(* IEC 61131-3 sources: llm-plc-st-eval/data/processed_v2/gpt-4o/I3/few_shot, 3 files *)

(* ---- ejec_1.st ---- *)
FUNCTION_BLOCK FB_Alarmas
VAR_INPUT
    alm1 : BOOL; (* Alarma 1 - Prioridad alta *)
    alm2 : BOOL; (* Alarma 2 - Prioridad media *)
    alm3 : BOOL; (* Alarma 3 - Prioridad baja *)
    ack1 : BOOL; (* Reconocimiento de alarma 1 *)
    ack2 : BOOL; (* Reconocimiento de alarma 2 *)
    ack3 : BOOL; (* Reconocimiento de alarma 3 *)
END_VAR
VAR_OUTPUT
    sirena : BOOL; (* Sirena de alarma *)
    codigoAlm : INT; (* Código de la alarma de mayor prioridad *)
END_VAR
VAR
    retAlm1 : BOOL; (* Retención de alarma 1 *)
    retAlm2 : BOOL; (* Retención de alarma 2 *)
    retAlm3 : BOOL; (* Retención de alarma 3 *)
END_VAR

(* Retención de alarmas *)
IF alm1 THEN
    retAlm1 := TRUE;
ELSIF ack1 AND NOT alm1 THEN
    retAlm1 := FALSE;
END_IF;

IF alm2 THEN
    retAlm2 := TRUE;
ELSIF ack2 AND NOT alm2 THEN
    retAlm2 := FALSE;
END_IF;

IF alm3 THEN
    retAlm3 := TRUE;
ELSIF ack3 AND NOT alm3 THEN
    retAlm3 := FALSE;
END_IF;

(* Determinación del código de alarma de mayor prioridad *)
IF retAlm1 THEN
    codigoAlm := 1;
ELSIF retAlm2 THEN
    codigoAlm := 2;
ELSIF retAlm3 THEN
    codigoAlm := 3;
ELSE
    codigoAlm := 0;
END_IF;

(* Activación de la sirena si hay cualquier alarma activa *)
sirena := retAlm1 OR retAlm2 OR retAlm3;

END_FUNCTION_BLOCK

(* ---- ejec_2.st ---- *)
FUNCTION_BLOCK FB_Alarmas
VAR_INPUT
    alm1 : BOOL; (* Alarma 1 - Alta prioridad *)
    alm2 : BOOL; (* Alarma 2 - Media prioridad *)
    alm3 : BOOL; (* Alarma 3 - Baja prioridad *)
    ack1 : BOOL; (* Reconocimiento de alarma 1 *)
    ack2 : BOOL; (* Reconocimiento de alarma 2 *)
    ack3 : BOOL; (* Reconocimiento de alarma 3 *)
END_VAR
VAR_OUTPUT
    sirena : BOOL; (* Sirena de alarma *)
    codigoAlm : INT; (* Código de alarma de mayor prioridad *)
END_VAR
VAR
    retAlm1 : BOOL; (* Retención de alarma 1 *)
    retAlm2 : BOOL; (* Retención de alarma 2 *)
    retAlm3 : BOOL; (* Retención de alarma 3 *)
END_VAR

(* Retención de alarmas *)
IF alm1 THEN
    retAlm1 := TRUE;
ELSIF ack1 AND NOT alm1 THEN
    retAlm1 := FALSE;
END_IF;

IF alm2 THEN
    retAlm2 := TRUE;
ELSIF ack2 AND NOT alm2 THEN
    retAlm2 := FALSE;
END_IF;

IF alm3 THEN
    retAlm3 := TRUE;
ELSIF ack3 AND NOT alm3 THEN
    retAlm3 := FALSE;
END_IF;

(* Determinación de la alarma de mayor prioridad *)
IF retAlm1 THEN
    codigoAlm := 1;
ELSIF retAlm2 THEN
    codigoAlm := 2;
ELSIF retAlm3 THEN
    codigoAlm := 3;
ELSE
    codigoAlm := 0;
END_IF;

(* Activación de la sirena si cualquier alarma está activa *)
sirena := retAlm1 OR retAlm2 OR retAlm3;
END_FUNCTION_BLOCK

(* ---- ejec_3.st ---- *)
FUNCTION_BLOCK FB_Alarmas
VAR_INPUT
    alm1 : BOOL; (* Alarma 1 - Alta prioridad *)
    alm2 : BOOL; (* Alarma 2 - Media prioridad *)
    alm3 : BOOL; (* Alarma 3 - Baja prioridad *)
    ack1 : BOOL; (* Reconocimiento de alarma 1 *)
    ack2 : BOOL; (* Reconocimiento de alarma 2 *)
    ack3 : BOOL; (* Reconocimiento de alarma 3 *)
END_VAR
VAR_OUTPUT
    sirena : BOOL; (* Sirena de alarma *)
    codigoAlm : INT; (* Código de alarma de mayor prioridad *)
END_VAR
VAR
    retAlm1 : BOOL; (* Retención de alarma 1 *)
    retAlm2 : BOOL; (* Retención de alarma 2 *)
    retAlm3 : BOOL; (* Retención de alarma 3 *)
END_VAR

(* Retención de alarmas *)
IF alm1 THEN
    retAlm1 := TRUE;
ELSIF ack1 AND NOT alm1 THEN
    retAlm1 := FALSE;
END_IF;

IF alm2 THEN
    retAlm2 := TRUE;
ELSIF ack2 AND NOT alm2 THEN
    retAlm2 := FALSE;
END_IF;

IF alm3 THEN
    retAlm3 := TRUE;
ELSIF ack3 AND NOT alm3 THEN
    retAlm3 := FALSE;
END_IF;

(* Determinación del código de alarma de mayor prioridad *)
IF retAlm1 THEN
    codigoAlm := 1;
ELSIF retAlm2 THEN
    codigoAlm := 2;
ELSIF retAlm3 THEN
    codigoAlm := 3;
ELSE
    codigoAlm := 0;
END_IF;

(* Activación de la sirena si hay alguna alarma retenida *)
sirena := retAlm1 OR retAlm2 OR retAlm3;

END_FUNCTION_BLOCK
